Fanuc KAREL source: kx00009.KL

-- PROVISIONAL review KL for V1013-1; original PC SHA256 8af250bf793ed0e2e240ba41fd4aca8af1d6b014a6d01297ee46e504597dc447
-- Incomplete behavior may be omitted. Consult companion uncertainty JSON. Do not deploy.
PROGRAM KX00009
%NOLOCKGROUP
VAR
  I : INTEGER
  J : INTEGER
  B : BOOLEAN
  F : FILE
  S : STRING[80]
-- UNRESOLVED_DECL P type=000102
BEGIN
  -- UNRESOLVED_PC offsets 5-7; opcodes 9C,4F
  -- UNRESOLVED_PC offsets 12-16; opcodes 7F
END KX00009
